(* IEC 61131-3 sources: ayran-mini-fabrika/plc/build (part 5) *)

  (* =================== 3. Shrink tunnel =================== *)
  (* if no new cup arrives for 2 minutes, energy saving; return to the normal setpoint when a new cup arrives *)
  T_IDLE(IN := MODE = 1 AND G_STP = 10 AND IW_LANE = LANE_LAST AND INSIDE = 0 AND W_STP = 0, PT := T#120s);
  LANE_LAST := IW_LANE;
  STANDBY := T_IDLE.Q;
  IF STANDBY THEN SP := SP_STANDBY; ELSE SP := SP_RUN; END_IF;
  TEMP_READY := (IW_TEMP >= SP_RUN - TEMP_BAND) AND (IW_TEMP <= SP_RUN + TEMP_BAND);

  (* outfeed blocked and packs in the tunnel: heater switches off immediately, packs are suspect *)
  T_EXITBLK(IN := DI_EXIT_FULL AND INSIDE > 0, PT := T#3s);
  IF T_EXITBLK.Q THEN HEAT_BLOCK := TRUE; END_IF;
  IF NOT DI_EXIT_FULL THEN HEAT_BLOCK := FALSE; END_IF;

  DRAINING := NOT WAIT_START AND MODE <> 1 AND MODE <> 4 AND INSIDE > 0 AND (ALARMS AND WORD#16#0180) = WORD#0;

  IF NOT ESTOP_OK OR NOT DI_FAN_RUN OR DI_OT_TRIP OR HEAT_BLOCK
     OR NOT (MODE = 1 OR DRAINING) OR (ALARMS AND WORD#16#00F0) <> WORD#0 THEN
    Q_HEAT := FALSE;
  ELSIF IW_TEMP < SP - HYST THEN
    Q_HEAT := TRUE;
  ELSIF IW_TEMP > SP + HYST THEN
    Q_HEAT := FALSE;
  END_IF;
  (* fan: does not stop while running, draining, or before the tunnel has cooled *)
  Q_FAN := NOT WAIT_START AND ESTOP_OK AND (MODE = 1 OR DRAINING OR IW_TEMP > COOL_OFF);
  Q_CONV := ESTOP_OK AND (MODE = 1 OR DRAINING) AND (ALARMS AND WORD#16#0080) = WORD#0;

  (* =================== 4. Grouping =================== *)
  T_PAD(IN := G_STP = 1, PT := T#3s);
  T_GATE(IN := G_STP = 11, PT := T#600ms);
  T_MOVE(IN := MODE = 1 AND NOT ROW_BLOCKED AND (G_STP = 12 OR G_STP = 13 OR G_STP = 21 OR G_STP = 22), PT := T#3s);

  IF MODE = 1 AND GROUP_OK THEN
    CASE G_STP OF
      0:  (* pad *)
        IF DI_ROWP_RET AND DI_GRPP_RET THEN
          IF ROWS >= 2 THEN G_STP := 20;
          ELSIF DI_PAD THEN G_STP := 10;
          ELSIF IW_PADS > 0 THEN G_STP := 1;
          END_IF;
        END_IF;
      1:
        IF DI_PAD THEN G_STP := 10; ELSIF T_PAD.Q THEN ALARMS := ALARMS OR WORD#16#0200; END_IF;
      10: (* let the lane fill *)
        IF ROWS >= 2 THEN G_STP := 20;
        ELSIF DI_LANE_FULL AND DI_ROWP_RET AND DI_GRPP_RET THEN G_STP := 11; END_IF;
      11: (* close the infeed gate, wait for the stroke *)
        IF T_GATE.Q THEN G_STP := 12; END_IF;
      12: (* row pusher forward *)
        IF DI_ROWP_EXT OR (ROWS >= 2 AND IW_LANE = 0) THEN G_STP := 13;
        ELSIF T_MOVE.Q THEN ALARMS := ALARMS OR WORD#16#0002; END_IF;
      13: (* back; a row is counted only when the pusher is back *)
        IF DI_ROWP_RET THEN
          IF ROWS >= 2 THEN G_STP := 20; ELSE G_STP := 10; END_IF;
        ELSIF T_MOVE.Q THEN
          ALARMS := ALARMS OR WORD#16#0002;
        END_IF;
      20: (* push the group when the wrapping machine is empty and ready *)
        IF ROWS = 0 THEN G_STP := 0;
        ELSIF ROWS >= 2 AND DI_WRAP_READY AND DI_ROWP_RET AND DI_GRPP_RET THEN G_STP := 21; END_IF;
      21:
        IF DI_GRPP_EXT THEN G_STP := 22; ELSIF T_MOVE.Q THEN ALARMS := ALARMS OR WORD#16#0004; END_IF;
      22:
        IF DI_GRPP_RET THEN G_STP := 0; ELSIF T_MOVE.Q THEN ALARMS := ALARMS OR WORD#16#0004; END_IF;
    END_CASE;
  END_IF;

  (* =================== 5. Wrapping and release =================== *)
  T_WRAP(IN := W_STP = 1, PT := T#6s);
  REL_OK := MODE = 1 AND TEMP_READY AND NOT STANDBY AND NOT DI_EXIT_FULL AND DI_BELT_RUN AND NOT HEAT_BLOCK;
  IF MODE = 1 THEN
    CASE W_STP OF
      0:
        IF DI_PACK_IN_WRAP THEN
          IF DI_WRAP_DONE THEN W_STP := 2; ELSE W_STP := 1; END_IF;
        END_IF;
      1:
        IF DI_WRAP_DONE THEN
          W_STP := 2;
        ELSIF T_WRAP.Q THEN
          ALARMS := ALARMS OR WORD#16#0008;
        END_IF;
      2:
        IF NOT DI_PACK_IN_WRAP THEN
          PACKS := PACKS + 1; IF PACKS > 30000 THEN PACKS := 0; END_IF;
          W_STP := 0;
        END_IF;
    END_CASE;
  END_IF;

  (* =================== 6. Outputs =================== *)
  Q_PAD  := MODE = 1 AND G_STP = 1;
  Q_GATE := G_STP >= 11 AND G_STP <= 13 AND MODE <> 4;
  Q_ROW  := MODE = 1 AND G_STP = 12 AND ROWS < 2;
  Q_GRP  := MODE = 1 AND G_STP = 21;
  Q_WRAP := MODE = 1 AND W_STP = 1;
  Q_REL  := W_STP = 2 AND REL_OK;

  QW_DO := WORD#0;
  IF Q_GATE THEN QW_DO := QW_DO OR WORD#16#0001; END_IF;
  IF Q_ROW  THEN QW_DO := QW_DO OR WORD#16#0002; END_IF;
  IF Q_GRP  THEN QW_DO := QW_DO OR WORD#16#0004; END_IF;
  IF Q_PAD  THEN QW_DO := QW_DO OR WORD#16#0008; END_IF;
  IF Q_WRAP THEN QW_DO := QW_DO OR WORD#16#0010; END_IF;
  IF Q_REL  THEN QW_DO := QW_DO OR WORD#16#0020; END_IF;
  IF Q_CONV THEN QW_DO := QW_DO OR WORD#16#0040; END_IF;
  IF Q_HEAT THEN QW_DO := QW_DO OR WORD#16#0080; END_IF;
  IF Q_FAN  THEN QW_DO := QW_DO OR WORD#16#0100; END_IF;
  IF Q_CONV AND NOT QUARANTINE THEN QW_DO := QW_DO OR WORD#16#0200; END_IF;
  IF Q_CONV AND QUARANTINE THEN QW_DO := QW_DO OR WORD#16#0400; END_IF;

  WARNS := WORD#0;
  IF HEAT_BLOCK THEN WARNS := WARNS OR WORD#16#0400; END_IF;
  IF IW_FILM < FILM_LOW THEN WARNS := WARNS OR WORD#16#0800; END_IF;
  IF DI_PAD_LOW THEN WARNS := WARNS OR WORD#16#1000; END_IF;
  QW_ALARM := ALARMS OR WARNS;

  (* state code and PackML-like status bits *)
  IF MODE = 4 THEN
    QW_STATE := 9;
  ELSIF MODE = 3 THEN
    IF DRAINING THEN QW_STATE := 5; ELSE QW_STATE := 8; END_IF;
  ELSIF MODE = 0 THEN
    IF DRAINING THEN
      QW_STATE := 5;
    ELSIF Q_FAN AND IW_TEMP > COOL_OFF THEN
      QW_STATE := 6;
    ELSE
      QW_STATE := 0;
    END_IF;
  ELSIF STANDBY THEN
    QW_STATE := 7;
  ELSIF NOT TEMP_READY THEN
    QW_STATE := 1;
  ELSIF W_STP = 2 AND NOT REL_OK AND DI_EXIT_FULL THEN
    QW_STATE := 4;
  ELSIF G_STP = 10 AND NOT DI_LANE_FULL THEN
    QW_STATE := 3;
  ELSE
    QW_STATE := 2;
  END_IF;

  STATUS := WORD#0;
  IF MODE = 1 AND G_STP = 10 THEN STATUS := STATUS OR WORD#16#0001; END_IF;
  IF MODE = 1 THEN STATUS := STATUS OR WORD#16#0002; END_IF;
  IF Q_HEAT AND NOT TEMP_READY THEN STATUS := STATUS OR WORD#16#0004; END_IF;
  IF DRAINING THEN STATUS := STATUS OR WORD#16#0008; END_IF;
  IF MODE = 3 OR MODE = 4 THEN STATUS := STATUS OR WORD#16#0010; END_IF;
  IF QW_STATE = 4 THEN STATUS := STATUS OR WORD#16#0020; END_IF;
  IF QW_STATE = 3 THEN STATUS := STATUS OR WORD#16#0040; END_IF;
  IF WAIT_START THEN STATUS := STATUS OR WORD#16#0080; END_IF;
  IF QUARANTINE THEN STATUS := STATUS OR WORD#16#0100; END_IF;
  QW_STATUS := STATUS;

  QW_PACKS  := PACKS;
  QW_INSIDE := INSIDE;
  QW_SP     := SP;
  QW_REJECT := IW_REJECT_CNT;
  QW_GOOD := IW_OUT_CNT - IW_REJECT_CNT;
  IF QW_GOOD < 0 THEN QW_GOOD := QW_GOOD + 30000; END_IF;
  RUNNING   := MODE = 1;
  IF WAIT_START OR NOT IO_READY THEN
    QW_DO := WORD#0;
    Q_HEAT := FALSE; Q_FAN := FALSE; Q_CONV := FALSE;
  END_IF;
END_FUNCTION_BLOCK

(* =====================================================================
   FB_Tank - tank, transfer line and CIP (block 2 of the factory)

   Line: sources V_PROD / V_WATER / V_CAUSTIC -> pump P1 -> flow meter FT1
        -> destinations V_FILL (filling tank) / V_DRAIN (drain) / V_CIPRET (caustic tank)

   Route manager: on every route change the pump stops, limit switches prove that
   all valves not in the new route are CLOSED, the new route
   is opened, the valve stroke time is waited out, and the pump starts again. If a valve not in
   the route appears open, the pump stops and an alarm is raised. This way caustic and
   product can never be in the same line at the same time.

   The filling machine requests product (REQ); this block transfers it or reports the reason it cannot.
   Times are at demo scale (in a real CIP the caustic contact time is 10-20 min).
   ===================================================================== *)

FUNCTION_BLOCK FB_Tank
  VAR_IN_OUT
    TNK_COMMISSION : WORD; (* one-shot commissioning token; consumed, never renewed by the FB *)
  END_VAR
  VAR_INPUT
    RESTART : BOOL;
    START : BOOL;
    ESTOP_OK, RESET : BOOL;   (* factory panel *)
    IO_READY   : BOOL;
    COMM_FAULT : BOOL;
    REQ        : BOOL;        (* the filling machine wants product *)
    IW_DI      : WORD;
    IW_T1_LVL  : INT;         (* 0.1 % *)
    IW_FLOW    : INT;         (* 0.01 kg/s *)
    IW_TOTAL   : INT;         (* 0.1 kg, wraps to zero at 30000 *)
    IW_COND    : INT;         (* 0.1 mS/cm, corrected to 25 C *)
    IW_RET_T   : INT;         (* 0.1 C *)
    IW_CIP_T   : INT;         (* 0.1 C *)
    IW_CIP_LVL : INT;         (* 0.1 % *)
  END_VAR
  VAR_OUTPUT
    QW_STATUS : WORD;
    QW_DO       : WORD;
    QW_STATE    : INT;
    QW_ALARM    : WORD;
    QW_STEP_T   : INT;
    QW_SINCE    : INT;
    QW_BATCH    : INT;
    QW_CIP_RES  : INT;
    QW_CIP_MINT : INT;
    QW_CIP_MINF : INT;
    QW_CIP_COND : INT;
    QW_CIP_DUR  : INT;
    TRANSFERRING : BOOL;
    CIP_DUE      : BOOL;
  END_VAR

  VAR
    (* ---- Recipe and settings (demo scale) ------------------------------ *)
    COND_MIN      : INT := 85;     (* product window 8.5..9.5 mS/cm (contains ~5% water) *)
    COND_MAX      : INT := 95;
    COND_CAUSTIC  : INT := 650;    (* effective caustic: >= 65 mS/cm (~80% concentration); sent to the return only at this concentration *)
    RINSE_MARGIN  : INT := 5;      (* final rinse: inlet water + 0.5 mS/cm *)
    FLOW_MIN      : INT := 50;     (* 0.5 kg/s *)
    FLOW_CIP      : INT := 150;    (* 1.5 kg/s for CIP *)
    CIP_TEMP_MIN  : INT := 700;    (* return temperature >= 70 C *)
    CAUSTIC_SP    : INT := 780;
    CAUSTIC_MAX   : INT := 900;
    CIP_LVL_MIN   : INT := 300;
    RINSE_KG      : INT := 300;    (* 30 kg of water per rinse *)
    CIP_LIMIT     : INT := 500;    (* one CIP per 50 kg of production *)
    ALARM_MASK    : WORD := WORD#16#23FF;   (* bits 0-9 and 13 are alarms, 10-12 are warnings *)
  END_VAR

  VAR
    (* ---- Decoded inputs ------------------------------------------- *)
    DI_T1_LOW, DI_CIP_START, DI_CIP_ABORT, DI_P1_RUN, DI_P1_TRIP, DI_LEAK : BOOL;
    CLOSED   : WORD;   (* aligned with the DO bits: bit1 V_PROD .. bit6 V_CIPRET *)

    (* ---- Route manager ---------------------------------------------- *)
    WANT     : WORD;   (* route requested by the step *)
    CUR      : WORD;   (* proven, applied route *)
    VALVES   : WORD;   (* command to the valves *)
    RSTATE       : INT;    (* 0 stable, 1 closing, 2 opening *)
    PUMP_REQ : BOOL;
    Q_P1     : BOOL;
    Q_HEAT   : BOOL;
    ROUTE_OK : BOOL;   (* all valves not in the route are closed *)

    (* ---- State -------------------------------------------------------- *)
    WAIT_START : BOOL := TRUE;
    MODE : INT := 0;
    RT_START : R_TRIG;
    STP        : INT := 0;
    LAST_STP   : INT := 0;
    STEP_SCANS  : INT;
    CIP_SCANS   : INT;
    ALARMS_BEFORE : WORD;
    ALARMS      : WORD;
    WARNS       : WORD;
    ABORT_WARN  : BOOL;
    LINE_PRODUCT : BOOL;   (* line is full of product and verified *)
    CIP_REQ     : BOOL;    (* the operator requested CIP; starts when the transfer ends *)
    CAUSTIC_IN  : BOOL;    (* caustic was routed to the return *)
    COND_OK     : BOOL;
    HOLD_OK     : BOOL;
    STEP_TO     : BOOL;
    TOTAL_LAST  : INT;
    TOTAL_INIT  : BOOL;
    D_TOTAL     : INT;
    SINCE       : INT;
    BATCH       : INT;
    VOL         : INT;
    WATER_REF   : INT;
    MIN_T       : INT;
    MIN_F       : INT;
    CIP_RES     : INT;
    FINAL_COND  : INT;
    CIP_DUR     : INT;

    (* ---- Timers (matiec: each on a separate line) --------------- *)
    RT_CIPSTART : R_TRIG;
    RT_CIPABORT : R_TRIG;
    RT_RESET    : R_TRIG;
    T_ROUTE     : TON;
    T_STROKE    : TON;
    T_LEAKVAL   : TON;
    T_NOFLOW    : TON;
    T_RUNFB     : TON;
    T_INWIN     : TON;
    T_FOREIGN   : TON;
    T_HOLD      : TON;
    T_STALE     : TON;
  END_VAR

  ALARMS_BEFORE := ALARMS;
  IF RESTART THEN
    MODE := 0; WAIT_START := TRUE;
    STP := 0; LAST_STP := 0; WANT := WORD#0; CUR := WORD#0; VALVES := WORD#0; RSTATE := 0;
    RSTATE := 1; (* prove all old-route valves closed *)
    Q_P1 := FALSE; Q_HEAT := FALSE; PUMP_REQ := FALSE; LINE_PRODUCT := FALSE; CIP_REQ := FALSE; TOTAL_INIT := FALSE;
    CIP_DUE := TNK_COMMISSION <> WORD#16#C1EA;
    IF CIP_DUE THEN CIP_RES := 2; ABORT_WARN := TRUE; END_IF;
    TNK_COMMISSION := WORD#0;
    T_ROUTE(IN := FALSE, PT := T#1s);
    T_STROKE(IN := FALSE, PT := T#1s);
    T_LEAKVAL(IN := FALSE, PT := T#1s);
    T_NOFLOW(IN := FALSE, PT := T#1s);
    T_RUNFB(IN := FALSE, PT := T#1s);
    T_INWIN(IN := FALSE, PT := T#1s);
    T_FOREIGN(IN := FALSE, PT := T#1s);
    T_HOLD(IN := FALSE, PT := T#1s);
    T_STALE(IN := FALSE, PT := T#1s);
  END_IF;

  (* =================== 1. Decode inputs =================== *)
  DI_T1_LOW    := (IW_DI AND WORD#16#0001) <> WORD#0;
  DI_CIP_START := (IW_DI AND WORD#16#0002) <> WORD#0;
  DI_CIP_ABORT := (IW_DI AND WORD#16#0004) <> WORD#0;
  DI_P1_RUN    := (IW_DI AND WORD#16#0008) <> WORD#0;
  DI_P1_TRIP   := (IW_DI AND WORD#16#0010) <> WORD#0;
  DI_LEAK      := (IW_DI AND WORD#16#0800) <> WORD#0;
  (* closed limit switches are DI bits 5..10; shifted right by 4 bits they align with DO bits 1..6 *)
  CLOSED := SHR(IW_DI, 4) AND WORD#16#007E;

  RT_CIPSTART(CLK := DI_CIP_START);
  RT_CIPABORT(CLK := DI_CIP_ABORT);
  RT_RESET(CLK := RESET);
  RT_START(CLK := START);
  IF RT_START.Q AND IO_READY AND NOT RESTART THEN WAIT_START := FALSE; MODE := 1; END_IF;

  (* increase of the flow meter totalizer in this scan (including wrap-around at 30000) *)
  IF NOT TOTAL_INIT THEN TOTAL_LAST := IW_TOTAL; TOTAL_INIT := IO_READY; END_IF;
  D_TOTAL := IW_TOTAL - TOTAL_LAST;
  IF D_TOTAL < 0 THEN D_TOTAL := D_TOTAL + 30000; END_IF;
  TOTAL_LAST := IW_TOTAL;

  COND_OK := (IW_COND >= COND_MIN) AND (IW_COND <= COND_MAX);

  (* =================== 2. Safety and alarms =================== *)
  IF NOT ESTOP_OK THEN ALARMS := ALARMS OR WORD#16#0001; END_IF;
  IF COMM_FAULT THEN ALARMS := ALARMS OR WORD#16#2000; END_IF;   (* no communication: stop safely *)
  IF DI_P1_TRIP THEN ALARMS := ALARMS OR WORD#16#0020; END_IF;
  IF DI_LEAK THEN ALARMS := ALARMS OR WORD#16#0010; END_IF;

  (* if a valve not in the route does not read closed for 1 s: valve stuck or leaking *)
  ROUTE_OK := ((NOT CUR) AND WORD#16#007E AND (NOT CLOSED)) = WORD#0;
  T_LEAKVAL(IN := RSTATE = 0 AND NOT ROUTE_OK, PT := T#1s);
  IF T_LEAKVAL.Q THEN ALARMS := ALARMS OR WORD#16#0008; END_IF;

  T_NOFLOW(IN := Q_P1 AND (IW_FLOW < FLOW_MIN), PT := T#3s);
  IF T_NOFLOW.Q THEN ALARMS := ALARMS OR WORD#16#0002; END_IF;
  T_RUNFB(IN := Q_P1 AND NOT DI_P1_RUN, PT := T#1s);
  IF T_RUNFB.Q THEN ALARMS := ALARMS OR WORD#16#0040; END_IF;

  IF IW_CIP_T > CAUSTIC_MAX THEN ALARMS := ALARMS OR WORD#16#0100; END_IF;

  IF NOT IO_READY THEN ALARMS := ALARMS_BEFORE; END_IF;

  (* alarm: everything shuts down; if a CIP is in progress it counts as failed *)
  IF (ALARMS AND ALARM_MASK) <> WORD#0 THEN
    IF STP >= 40 THEN CIP_RES := 3; CIP_DUE := TRUE; LINE_PRODUCT := FALSE; END_IF;
    STP := 0;
  END_IF;

  IF RT_RESET.Q THEN
    IF ESTOP_OK AND NOT COMM_FAULT AND NOT DI_P1_TRIP AND NOT DI_LEAK THEN
      ALARMS := WORD#0;
    END_IF;
  END_IF;

  (* =================== 3. Steps =================== *)
  (* note: STEP and RS are IEC 61131-3 reserved words (SFC step, RS flip-flop); STP / RSTATE are used instead *)
  IF STP <> LAST_STP THEN STEP_SCANS := 0; VOL := 0; END_IF;
  LAST_STP := STP;
  IF STEP_SCANS < 30000 THEN STEP_SCANS := STEP_SCANS + 1; END_IF;
  IF RSTATE = 0 AND (STP = 42 OR STP = 44) THEN VOL := VOL + D_TOTAL; END_IF;

  (* quantity passed through the route applied for production *)
  IF CUR = WORD#16#0012 OR CUR = WORD#16#0022 THEN
    IF SINCE < 30000 THEN SINCE := SINCE + D_TOTAL; END_IF;
  END_IF;
  IF CUR = WORD#16#0012 THEN BATCH := BATCH + D_TOTAL; END_IF;
  IF SINCE >= CIP_LIMIT THEN CIP_DUE := TRUE; END_IF;

  (* product waiting in the line for a long time goes stale: a push-out is needed again *)
  T_STALE(IN := STP = 0 AND LINE_PRODUCT, PT := T#1200s);
  IF T_STALE.Q THEN LINE_PRODUCT := FALSE; END_IF;

  IF RT_CIPSTART.Q THEN CIP_REQ := TRUE; END_IF;

  (* CIP abort *)
  IF RT_CIPABORT.Q AND STP >= 40 THEN
    CIP_RES := 2;
    CIP_DUE := TRUE;
    CIP_REQ := FALSE;
    ABORT_WARN := TRUE;
    LINE_PRODUCT := FALSE;
    STP := 0;
  END_IF;

  T_INWIN(IN := STP = 20 AND RSTATE = 0 AND Q_P1 AND COND_OK, PT := T#1s);
  T_FOREIGN(IN := STP = 10 AND RSTATE = 0 AND Q_P1 AND NOT COND_OK, PT := T#1s);
  HOLD_OK := STP = 43 AND RSTATE = 0 AND CUR = WORD#16#0048 AND Q_P1
             AND IW_COND >= COND_CAUSTIC AND IW_RET_T >= CIP_TEMP_MIN AND IW_FLOW >= FLOW_CIP;
  T_HOLD(IN := HOLD_OK, PT := T#30s);
  STEP_TO := STEP_SCANS >= 15000;     (* 300 s; with a 20 ms task cycle *)

  CASE STP OF
    0:  (* idle *)
      WANT := WORD#0;
      PUMP_REQ := FALSE;
      IF NOT WAIT_START AND (ALARMS AND ALARM_MASK) = WORD#0 THEN
        IF CIP_REQ THEN
          CIP_REQ := FALSE;
          STP := 40;
        ELSIF REQ AND NOT CIP_DUE AND NOT DI_T1_LOW THEN
          BATCH := 0;
          IF LINE_PRODUCT THEN STP := 10; ELSE STP := 20; END_IF;
        END_IF;
      END_IF;

    20: (* fill the line with product: first liquid to the drain *)
      WANT := WORD#16#0022;            (* V_PROD + V_DRAIN *)
      PUMP_REQ := TRUE;
      IF T_INWIN.Q THEN
        LINE_PRODUCT := TRUE;
        STP := 10;                     (* the route manager stops the pump and changes the route *)
      ELSIF STEP_SCANS > 2250 THEN
        ALARMS := ALARMS OR WORD#16#0200;   (* product conductivity not detected within 45 s *)
      END_IF;

    10: (* transfer to the filling tank *)
      WANT := WORD#16#0012;            (* V_PROD + V_FILL *)
      PUMP_REQ := TRUE;
      IF T_FOREIGN.Q THEN
        LINE_PRODUCT := FALSE;
        ALARMS := ALARMS OR WORD#16#0004;
      ELSIF NOT REQ OR DI_T1_LOW OR SINCE >= CIP_LIMIT OR CIP_REQ THEN
        STP := 0;
      END_IF;

    40: (* CIP preparation: empty route for the line, prove all valves closed *)
      WANT := WORD#0;
      PUMP_REQ := FALSE;
      LINE_PRODUCT := FALSE;
      CAUSTIC_IN := FALSE;
      CIP_SCANS := 0;
      MIN_T := 32000;
      MIN_F := 32000;
      FINAL_COND := 0;
      IF IW_CIP_LVL < CIP_LVL_MIN THEN
        ALARMS := ALARMS OR WORD#16#0100;
      ELSIF RSTATE = 0 AND ROUTE_OK THEN
        STP := 41;
      END_IF;

    41: (* wait for the caustic temperature *)
      WANT := WORD#0;
      PUMP_REQ := FALSE;
      IF IW_CIP_T >= CAUSTIC_SP - 50 THEN
        STP := 42;
      ELSIF STEP_TO THEN
        ALARMS := ALARMS OR WORD#16#0080;
      END_IF;

    42: (* pre-rinse: water to the drain *)
      WANT := WORD#16#0024;            (* V_WATER + V_DRAIN *)
      PUMP_REQ := TRUE;
      IF VOL >= RINSE_KG THEN
        WATER_REF := IW_COND;           (* conductivity of the inlet water: the criterion for the final rinse *)
        STP := 43;
      ELSIF STEP_TO THEN
        ALARMS := ALARMS OR WORD#16#0080;
      END_IF;

    43: (* caustic: first to the drain, to the caustic tank once caustic arrives (phase separation) *)
      PUMP_REQ := TRUE;
      IF NOT CAUSTIC_IN AND RSTATE = 0 AND IW_COND >= COND_CAUSTIC THEN CAUSTIC_IN := TRUE; END_IF;
      IF CAUSTIC_IN THEN
        WANT := WORD#16#0048;          (* V_CAUSTIC + V_CIPRET *)
      ELSE
        WANT := WORD#16#0028;          (* V_CAUSTIC + V_DRAIN *)
      END_IF;
      (* CIP record: the lowest values in the counted hold window *)
      IF HOLD_OK THEN
        IF IW_RET_T < MIN_T THEN MIN_T := IW_RET_T; END_IF;
        IF IW_FLOW < MIN_F THEN MIN_F := IW_FLOW; END_IF;
      ELSE
        MIN_T := 32000;
        MIN_F := 32000;
      END_IF;
      IF T_HOLD.Q THEN
        STP := 44;
      ELSIF STEP_TO THEN
        ALARMS := ALARMS OR WORD#16#0080;
      END_IF;

    44: (* final rinse: until no caustic is left *)
      WANT := WORD#16#0024;
      PUMP_REQ := TRUE;
      IF VOL >= RINSE_KG AND IW_COND <= WATER_REF + RINSE_MARGIN THEN
        FINAL_COND := IW_COND;
        STP := 45;
      ELSIF STEP_TO THEN
        ALARMS := ALARMS OR WORD#16#0080;
      END_IF;

    45: (* completed *)
      WANT := WORD#0;
      PUMP_REQ := FALSE;
      SINCE := 0;
      CIP_DUE := FALSE;
      ABORT_WARN := FALSE;
      CIP_RES := 1;
      CIP_DUR := CIP_SCANS / 50;
      STP := 0;
  END_CASE;
  IF STP >= 40 AND STP <= 44 AND CIP_SCANS < 30000 THEN CIP_SCANS := CIP_SCANS + 1; END_IF;
  IF CIP_RES = 2 OR CIP_RES = 3 THEN CIP_DUR := CIP_SCANS / 50; END_IF;

  (* =================== 4. Route manager =================== *)
  IF (ALARMS AND ALARM_MASK) <> WORD#0 THEN WANT := WORD#0; END_IF;
  IF WANT <> CUR AND RSTATE = 0 THEN RSTATE := 1; END_IF;
  T_ROUTE(IN := RSTATE = 1, PT := T#3s);
  T_STROKE(IN := RSTATE = 2, PT := T#1s);
  IF RSTATE = 1 THEN
    VALVES := CUR AND WANT;            (* close the ones not in the new route *)
    IF ((NOT WANT) AND WORD#16#007E AND (NOT CLOSED)) = WORD#0 THEN
      RSTATE := 2;
    ELSIF T_ROUTE.Q THEN
      ALARMS := ALARMS OR WORD#16#0008;
      RSTATE := 0;
      CUR := CUR AND WANT;
    END_IF;
  ELSIF RSTATE = 2 THEN
    VALVES := WANT;
    IF T_STROKE.Q THEN CUR := WANT; RSTATE := 0; END_IF;
  ELSE
    VALVES := CUR;
  END_IF;

  Q_P1 := PUMP_REQ AND RSTATE = 0 AND CUR = WANT AND CUR <> WORD#0 AND ROUTE_OK
          AND (ALARMS AND ALARM_MASK) = WORD#0;

  (* caustic tank thermostat (+/- 2 C), level and over-temperature interlock *)
  IF NOT ESTOP_OK OR IW_CIP_LVL < CIP_LVL_MIN OR IW_CIP_T > CAUSTIC_MAX THEN
    Q_HEAT := FALSE;
  ELSIF IW_CIP_T < CAUSTIC_SP - 20 THEN
    Q_HEAT := TRUE;
  ELSIF IW_CIP_T > CAUSTIC_SP + 20 THEN
    Q_HEAT := FALSE;
  END_IF;

  (* =================== 5. Outputs =================== *)
  WARNS := WORD#0;
  IF DI_T1_LOW THEN WARNS := WARNS OR WORD#16#0400; END_IF;
  IF CIP_DUE THEN WARNS := WARNS OR WORD#16#0800; END_IF;
  IF ABORT_WARN THEN WARNS := WARNS OR WORD#16#1000; END_IF;

  QW_DO := VALVES AND WORD#16#007E;
  IF Q_P1 THEN QW_DO := QW_DO OR WORD#16#0001; END_IF;
  IF Q_HEAT THEN QW_DO := QW_DO OR WORD#16#0080; END_IF;
  IF STP >= 40 THEN QW_DO := QW_DO OR WORD#16#0100; END_IF;

  IF (ALARMS AND WORD#16#0001) <> WORD#0 THEN
    QW_STATE := 11;
  ELSIF (ALARMS AND ALARM_MASK) <> WORD#0 THEN
    QW_STATE := 10;
  ELSIF STP = 0 AND CIP_DUE THEN
    QW_STATE := 9;
  ELSIF STP = 0 THEN
    QW_STATE := 0;
  ELSIF (STP = 10 OR STP = 20) AND RSTATE <> 0 THEN
    QW_STATE := 3;
  ELSIF STP = 10 THEN
    QW_STATE := 1;
  ELSIF STP = 20 THEN
    QW_STATE := 2;
  ELSE
    QW_STATE := STP - 36;             (* 40..44 -> 4..8 *)
  END_IF;

  QW_ALARM    := ALARMS OR WARNS;
  QW_STEP_T   := STEP_SCANS / 50;
  QW_SINCE    := SINCE;
  QW_BATCH    := BATCH;
  QW_CIP_RES  := CIP_RES;
  IF MIN_T = 32000 THEN QW_CIP_MINT := 0; ELSE QW_CIP_MINT := MIN_T; END_IF;
  IF MIN_F = 32000 THEN QW_CIP_MINF := 0; ELSE QW_CIP_MINF := MIN_F; END_IF;
  QW_CIP_COND := FINAL_COND;
  QW_CIP_DUR  := CIP_DUR;
  TRANSFERRING := STP = 10 AND Q_P1;
  QW_STATUS := WORD#0;
  IF WAIT_START THEN QW_STATUS := WORD#16#0080; END_IF;
  IF WAIT_START OR NOT IO_READY THEN
    QW_DO := WORD#0;
    Q_HEAT := FALSE; Q_P1 := FALSE;
  END_IF;
END_FUNCTION_BLOCK

PROGRAM Paketleme
  VAR
    (* --- blok 0: Fabrika --- *)
    FAB_IW_DI        AT %IW100 : WORD;  (* Fabrika paneli girisleri (bit paketli) *)
    FAB_IW_MAPVER    AT %IW101 : INT;  (* Sinyal haritasi surumu *)
    FAB_IW_SIM_HB    AT %IW102 : INT;  (* Simulator kalp atisi (100 ms) *)
    (* --- blok 1: Dolum-kapama --- *)
    DOL_IW_DI        AT %IW116 : WORD;  (* Dijital girisler (bit paketli) *)
    DOL_IW_FILL      AT %IW117 : INT;  (* Dolum terazisi (net) *)
    DOL_IW_TANK      AT %IW118 : INT;  (* Dolum tanki seviyesi *)
    DOL_IW_TEMP      AT %IW119 : INT;  (* Kapama kafasi sicakligi *)
    DOL_IW_CHECK     AT %IW120 : INT;  (* Kontrol tartisi (brut) *)
    (* --- blok 2: Tank ve transfer --- *)
    TNK_IW_DI        AT %IW132 : WORD;  (* Dijital girisler (bit paketli) *)
    TNK_IW_T1_LVL    AT %IW133 : INT;  (* Uretim tanki T1 seviyesi *)
    TNK_IW_FLOW      AT %IW134 : INT;  (* Debimetre FT1 *)
    TNK_IW_TOTAL     AT %IW135 : INT;  (* Debimetre toplayici (30000'de sifirlanir) *)
    TNK_IW_COND      AT %IW136 : INT;  (* Hat iletkenligi QT1 (25 ?C'ye duzeltilmis) *)
    TNK_IW_RET_T     AT %IW137 : INT;  (* Hat donus sicakligi TT1 *)
    TNK_IW_CIP_T     AT %IW138 : INT;  (* Kostik tanki sicakligi TT2 *)
    TNK_IW_CIP_LVL   AT %IW139 : INT;  (* Kostik tanki seviyesi *)
    (* --- blok 3: Shrink ve firin --- *)
    SHR_IW_DI        AT %IW148 : WORD;  (* Dijital girisler (bit paketli) *)
    SHR_IW_LANE      AT %IW149 : INT;  (* Seritteki bardak sayisi (bilesik sensor) *)
    SHR_IW_TEMP      AT %IW150 : INT;  (* Firin hava sicakligi *)
    SHR_IW_IN_CNT    AT %IW151 : INT;  (* Firin girisi paket sayaci (30000'de sifirlanir) *)
    SHR_IW_OUT_CNT   AT %IW152 : INT;  (* Firin cikisi paket sayaci *)
    SHR_IW_FILM      AT %IW153 : INT;  (* Film bobini kalan *)
    SHR_IW_PADS      AT %IW154 : INT;  (* Altlik magazini adedi *)
    SHR_IW_EXIT_CNT  AT %IW155 : INT;  (* Cikistan alinan paket sayaci *)
    SHR_IW_PLATE     AT %IW156 : WORD;  (* Plaka fotoselleri (bit 0: sira 1, bit 1: sira 2) *)
    SHR_IW_DIVERT    AT %IW157 : WORD;  (* Cikis ayirici: bit 0 paket var, 1 red konumu, 2 gecis konumu *)
    SHR_IW_REJECT_CNT AT %IW158 : INT;  (* Karantina kasasina ayrilan paket sayaci (30000 modul) *)
    SHR_QW_DO        AT %QW100 : WORD;  (* Dijital cikislar (bit paketli) *)
    SHR_QW_STATE     AT %QW101 : INT;  (* Istasyon durumu *)
    SHR_QW_ALARM     AT %QW102 : WORD;  (* Alarm kelimesi *)
    SHR_QW_STATUS    AT %QW103 : WORD;  (* Durum bitleri (PackML benzeri) *)
    SHR_QW_PACKS     AT %QW104 : INT;  (* Firina birakilan paket sayaci *)
    SHR_QW_INSIDE    AT %QW105 : INT;  (* Firin icindeki paket *)
    SHR_QW_SP        AT %QW106 : INT;  (* Gecerli firin ayar degeri *)
    SHR_QW_REJECT    AT %QW107 : INT;  (* Fotoselden dogrulanan karantina paket sayaci (30000 modul) *)
    SHR_QW_GOOD      AT %QW108 : INT;  (* Iyi urun bandina gecirilen paket sayaci (30000 modul) *)
    SHR_QW_PLC_HB    AT %QW115 : INT;  (* Paketleme PLC kalp atisi (her tarama) *)
    (* --- blok 4: Paletleme --- *)
    PAL_IW_DI        AT %IW164 : WORD;  (* Hat ve guvenlik girisleri (bit paketli) *)
    PAL_IW_ROB_DI    AT %IW165 : WORD;  (* Robot kontrolcusu durum bitleri *)
    PAL_IW_ACK_SEQ   AT %IW166 : INT;  (* Robot: kabul edilen son is numarasi *)
    PAL_IW_RES_SEQ   AT %IW167 : INT;  (* Robot: biten son is numarasi *)
    PAL_IW_RES_CODE  AT %IW168 : INT;  (* Robot: son is sonucu (1 tamam, 10+ hata) *)
    PAL_IW_RES_SLOT  AT %IW169 : INT;  (* Robot: son isin slotu *)
    PAL_IW_TURNS     AT %IW170 : INT;  (* Strec sarma: bu cevrimdeki tur *)
    PAL_IW_PALLETS   AT %IW171 : INT;  (* Bos palet magazini adedi *)
    PAL_IW_SHEETS    AT %IW172 : INT;  (* Karton levha magazini adedi *)
    PAL_IW_PICKUP_CNT AT %IW173 : INT;  (* Alim noktasindan alinan palet sayaci *)
    PAL_IW_IL        AT %IW174 : WORD;  (* Istasyon el sikisma girisleri (AGV optik I/O) *)
    PAL_IW_RES_JOB   AT %IW175 : INT;  (* Robot: biten son isin tipi *)
    PAL_QW_DO        AT %QW116 : WORD;  (* Dijital cikislar (bit paketli) *)
    PAL_QW_JOB       AT %QW117 : INT;  (* Robot isi (1 al, 2 birak, 3 levha, 4 eve don) *)
    PAL_QW_SLOT      AT %QW118 : INT;  (* Robot slotu (birak: 1..18, levha: 0 alt / 1 ust) *)
    PAL_QW_SEQ       AT %QW119 : INT;  (* Robot is numarasi (degisince is baslar) *)
    PAL_QW_STATE     AT %QW120 : INT;  (* Istasyon durumu *)
    PAL_QW_ALARM     AT %QW121 : WORD;  (* Alarm kelimesi *)
    PAL_QW_STATUS    AT %QW122 : WORD;  (* Durum bitleri (PackML benzeri) *)
    PAL_QW_COUNT     AT %QW123 : INT;  (* Istifteki paletin paket sayisi (dogrulanmis) *)
    PAL_QW_DONE      AT %QW124 : INT;  (* Tamamlanan palet sayaci *)
    PAL_QW_PALLET_ID AT %QW125 : INT;  (* Istifteki paletin numarasi *)
    PAL_QW_WRAPPED   AT %QW126 : INT;  (* Streclenen palet sayaci *)
    RET_MAGIC AT %MW32 : WORD;
    RET_MAPVER AT %MW33 : INT;
    PAL_COUNT AT %MW34 : INT;
    PAL_ID AT %MW35 : INT;
    PAL_DONE AT %MW36 : INT;
    PAL_WRAPPED AT %MW37 : INT;
    PAL_SHEETS AT %MW38 : WORD;
    PAL_LAST_SEQ AT %MW39 : INT;
    PAL_ACTIVE AT %MW40 : WORD;
    PAL_C_PHASE AT %MW41 : INT;
    PAL_UNDERWRAP AT %MW42 : WORD;
    RET_CHECK AT %MW43 : WORD;
  END_VAR

  VAR
    PB_START    : BOOL;   (* factory panel *)
    PB_STOP_OK  : BOOL;
    PB_ESTOP_OK : BOOL;
    PB_RESET    : BOOL;
    FIRST_SCAN  : BOOL := TRUE;
    RESTART     : BOOL;
    IO_READY    : BOOL;   (* first data arrived from the simulator with the correct version *)
    COMM_FAULT  : BOOL;
    SIM_HB_LAST : INT;
    PLC_HB      : INT;
    T_SIMHB     : TON;
    SHRINK      : FB_Shrink;
    PALLET      : FB_Pallet;
  END_VAR

  (* =================== 1. Factory panel =================== *)
  PB_START    := (FAB_IW_DI AND WORD#16#0001) <> WORD#0;
  PB_STOP_OK  := (FAB_IW_DI AND WORD#16#0002) <> WORD#0;
  PB_ESTOP_OK := (FAB_IW_DI AND WORD#16#0004) <> WORD#0;
  PB_RESET    := (FAB_IW_DI AND WORD#16#0008) <> WORD#0;

  (* =================== 2. Communication watchdog =================== *)
  (* communication fault if the simulator heartbeat does not change for 2 s *)
  T_SIMHB(IN := (FAB_IW_SIM_HB = SIM_HB_LAST), PT := T#2s);
  SIM_HB_LAST := FAB_IW_SIM_HB;
  COMM_FAULT := T_SIMHB.Q;
  (* inputs are invalid until the first data arrives and the map version matches *)
  IF FAB_IW_SIM_HB <> 0 AND FAB_IW_MAPVER = 7 THEN IO_READY := TRUE; END_IF;

  RESTART := FIRST_SCAN AND IO_READY;
  IF RESTART THEN FIRST_SCAN := FALSE; END_IF;

  (* PLC heartbeat: the simulator watches it and switches off this PLC's outputs if the program stops *)
  PLC_HB := PLC_HB + 1;
  IF PLC_HB > 30000 THEN PLC_HB := 0; END_IF;

  (* =================== Grouping, wrapping, shrink tunnel =================== *)
  (* contract: when the outfeed belt is full the filler already waits, and this station in turn
     releases no pack into the tunnel when its own outfeed is full *)
  SHRINK(START := PB_START, STOP_OK := PB_STOP_OK, ESTOP_OK := PB_ESTOP_OK, RESET := PB_RESET,
         RESTART := RESTART, IO_READY := IO_READY, COMM_FAULT := COMM_FAULT,
         IW_DI := SHR_IW_DI, IW_LANE := SHR_IW_LANE, IW_TEMP := SHR_IW_TEMP,
         IW_IN_CNT := SHR_IW_IN_CNT, IW_OUT_CNT := SHR_IW_OUT_CNT, IW_FILM := SHR_IW_FILM, IW_PADS := SHR_IW_PADS,
         IW_PLATE := SHR_IW_PLATE, IW_REJECT_CNT := SHR_IW_REJECT_CNT);
  SHR_QW_DO     := SHRINK.QW_DO;
  SHR_QW_STATE  := SHRINK.QW_STATE;
  SHR_QW_ALARM  := SHRINK.QW_ALARM;
  SHR_QW_STATUS := SHRINK.QW_STATUS;
  SHR_QW_PACKS  := SHRINK.QW_PACKS;
  SHR_QW_INSIDE := SHRINK.QW_INSIDE;
  SHR_QW_SP     := SHRINK.QW_SP;
  SHR_QW_REJECT := SHRINK.QW_REJECT;
  SHR_QW_GOOD := SHRINK.QW_GOOD;

  (* =================== Robotic palletizing =================== *)
  (* contract: if the robot does not take the pack at the pickup point, the tunnel outfeed fills up and
     the shrink tunnel accepts no new pack. The AGV's "forks outside the pickup point" signal is the
     optical signal the vehicle gives to the station: the station's own input (PAL_IW_IL bit 0); it
     does not pass through the logistics PLC. *)
  PALLET(START := PB_START, STOP_OK := PB_STOP_OK, ESTOP_OK := PB_ESTOP_OK, RESET := PB_RESET,
         RESTART := RESTART, IO_READY := IO_READY, COMM_FAULT := COMM_FAULT,
         IW_DI := PAL_IW_DI, IW_ROB_DI := PAL_IW_ROB_DI, IW_ACK_SEQ := PAL_IW_ACK_SEQ, IW_RES_SEQ := PAL_IW_RES_SEQ,
         IW_RES_JOB := PAL_IW_RES_JOB, IW_RES_CODE := PAL_IW_RES_CODE, IW_RES_SLOT := PAL_IW_RES_SLOT, IW_TURNS := PAL_IW_TURNS,
         IW_PALLETS := PAL_IW_PALLETS, IW_SHEETS := PAL_IW_SHEETS,
         AGV_CLEAR := (PAL_IW_IL AND WORD#16#0001) <> WORD#0,
         RET_MAGIC := RET_MAGIC, RET_MAPVER := RET_MAPVER, PAL_COUNT := PAL_COUNT, PAL_ID := PAL_ID,
         PAL_DONE := PAL_DONE, PAL_WRAPPED := PAL_WRAPPED, PAL_SHEETS := PAL_SHEETS,
         PAL_LAST_SEQ := PAL_LAST_SEQ, PAL_ACTIVE := PAL_ACTIVE, PAL_C_PHASE := PAL_C_PHASE,
         PAL_UNDERWRAP := PAL_UNDERWRAP, RET_CHECK := RET_CHECK);
  PAL_QW_DO        := PALLET.QW_DO;
  PAL_QW_JOB       := PALLET.QW_JOB;
  PAL_QW_SLOT      := PALLET.QW_SLOT;
  PAL_QW_SEQ       := PALLET.QW_SEQ;
  PAL_QW_STATE     := PALLET.QW_STATE;
  PAL_QW_ALARM     := PALLET.QW_ALARM;
  PAL_QW_STATUS    := PALLET.QW_STATUS;
  PAL_QW_COUNT     := PALLET.QW_COUNT;
  PAL_QW_DONE      := PALLET.QW_DONE;
  PAL_QW_PALLET_ID := PALLET.QW_PALLET_ID;
  PAL_QW_WRAPPED   := PALLET.QW_WRAPPED;

  SHR_QW_PLC_HB := PLC_HB;
END_PROGRAM

CONFIGURATION Config0
  RESOURCE Res0 ON PLC
    TASK task0(INTERVAL := T#20ms, PRIORITY := 0);
    PROGRAM instance0 WITH task0 : Paketleme;
  END_RESOURCE
END_CONFIGURATION
